Fanuc KAREL source: KT00740.KL

PROGRAM KT00740
%NOLOCKGROUP
VAR
  ARG: ARRAY[4] OF SHORT
  OUT: BOOLEAN
BEGIN
  OUT = UNINIT(ARG)
END KT00740
